PROGRAM MAIN
VAR
	fb_Startup : FB_Startup;
	fb_ModbusComm: FB_ModbusComm;
	fb_System_Time : FB_System_Time;
	fb_Jog_Joint : FB_Jog_Joint;
	fb_ElectromagnetActivate : FB_ElectromagnetActivate;
END_VAR


(*
GJENSTÅENDE ARBEID:
1) Implementer auto sekvens FB
2) 
*)


GVL.LED_J1_CW := GVL.PB_J1_CW;
GVL.LED_J2_CW := GVL.PB_J2_CW;
GVL.LED_J3_CW := GVL.PB_J3_CW;
GVL.LED_J1_CCW := GVL.PB_J1_CCW;
GVL.LED_J2_CCW := GVL.PB_J2_CCW;
GVL.LED_J3_CCW := GVL.PB_J3_CCW;
GVL.LED_EE_Grip := GVL.PB_EE_Grip;
GVL.LED_EE_Ungrip := GVL.PB_EE_Ungrip;
GVL.LED_EMG_STOP := NOT GVL.PB_EMG_STOP;
GVL.LED_Start_Pause := GVL.PB_Start_Pause;
GVL.LED_Reset := GVL.LED_Reset;
GVL.LED_Warning := TRUE;
GVL.LED_Reset := GVL.PB_Reset;
GVL.LED_Start_Pause := GVL.PB_Start_Pause;
GVL.LED_Record_Pos := GVL.PB_Record_Pos;


// Code which must run every PLC cycle.
fb_System_Time(); // Run FB to calculate Delta_Time


(* COMMENTING OUT FOR TESTING PURPOSES
IF NOT GVL.PB_EMG_STOP AND NOT (gvl.system_state = state_enum.startup_mode) THEN
	GVL.system_state := state_enum.emg_stop_mode;
ELSIF GVL.LED_Comm_Fault AND NOT (gvl.system_state = state_enum.startup_mode)  THEN
	GVL.system_state := state_enum.comm_fault_mode;
END_IF
*)


CASE gvl.system_state OF
state_enum.startup_mode:
	fb_Startup();
state_enum.jog_joint_mode:
	fb_Jog_Joint(
	lr_DeltaTime:= fb_ModbusComm.lreal_CycleTime, 
	lr_SlowModeVelocitySetting:= 1, 
	lr_FastModeVelovitySetting:= 10, 
	i_Base_LowLimit:= 0, 
	i_Base_HighLimit:= 180, 
	i_Shoulder_LowLimit:= 0, 
	i_Shoulder_HighLimit:= 180, 
	i_Elbow_LowLimit:= 0, 
	i_Elbow_HighLimit:= 180, 
	b_Enable_Servos:= TRUE, 
	SW_Fast_Mode:= GVL.SW_Slow_Fast, 
	PB_Base_Pos:= GVL.PB_J1_CCW, 
	PB_Base_Neg:= GVL.PB_J1_CW, 
	PB_Shoulder_Pos:= GVL.PB_J2_CCW, 
	PB_Shoulder_Neg:= GVL.PB_J2_CW, 
	PB_Elbow_Pos:= GVL.PB_J3_CCW, 
	PB_Elbow_Neg:= GVL.PB_J3_CW, 
	i_Set_Base=>, 
	i_Set_Shoulder=>, 
	i_Set_Elbow=>);
	
	fb_ElectromagnetActivate(
	b_activate := GVL.PB_EE_Grip,
	b_deactivate := GVL.PB_EE_Ungrip,
	b_CMD_Magnet =>);
	
state_enum.jog_cartesian_mode:
state_enum.manual_mode:
state_enum.emg_stop_mode:
state_enum.comm_fault_mode:
state_enum.auto_mode:
END_CASE

//fb_ModbusComm();
fb_ModbusComm(
	i_MBO_BaseAngle:= fb_Jog_Joint.i_Set_Base, 
	i_MBO_ShoulderAngle:= fb_Jog_Joint.i_Set_Shoulder, 
	i_MBO_ElbowAngle:= fb_Jog_Joint.i_Set_Elbow, 
	i_MBO_EndEffectorValue:= BOOL_TO_INT(fb_ElectromagnetActivate.b_CMD_Magnet), 
	b_MBO_EmergencyStop:= , 
	lreal_CycleTime := fb_System_Time.Delta_Time,
	iLastWrittenBaseAngle=> , 
	iLastWrittenShoulderAngle=> , 
	iLastWrittenElbowAngle=> , 
	b_MBI_LocalControl=> , 
	b_MBI_LocalEmergencyStopActive=> , 
	b_MBWatchdogTimeout=> GVL.LED_Comm_Fault, 
	i_MBI_LocalBaseAngle=> , 
	i_MBI_LocalShoulderAngle=> , 
	i_MBI_LocalElbowAngle=> , 
	i_MBI_LocalValueEndEffector=> );

END_PROGRAM

(* stored: Version 1.1.0.1, ProductVersion 3.1.4024.13
   POU MAIN: Id {5c661849-addd-4c08-be03-d943d6f2eed1}, SpecialFunc None *)
